Staubli VAL3: click_refreshTrajMsg.pgx

program click_refreshTrajMsg()
begin
  nMsgType=2
  call initMsg()
  call rs:getLog(sRobotMsg,nMsgType)
  userPageSet("message","btnAllMsg","style.backgroundColor","#FFFFFF")
  userPageSet("message","btnRobotMsg","style.backgroundColor","#FFFFFF")
  userPageSet("message","btnTrajMsg","style.backgroundColor","#33FF33")
  userPageSet("message","btnIOMsg","style.backgroundColor","#FFFFFF")
end
